% RSLogix 500 project MIXING.RSS, saved by version 8.30.00.16 %
PROJECT "UNTITLED"    % processor: MicroLogix 1000 %

PROGRAM FILES
  LAD 2 "MAIN_PROG"  6 rungs
  LAD 3 "USER_FAULT"  1 rungs
  LAD 4 "HSC_INT"  1 rungs
  LAD 5 "STI_INT"  1 rungs
  LAD 6, 7, 8, 9, 10, 11, 12, 13, 14, 15, 16: only END

DATA FILES
  O0 OUTPUT  5 elements
  I1 INPUT  8 elements
  S2 STATUS  33 elements
  B3 BINARY  32 elements
  T4 TIMER  40 elements
  C5 COUNTER  32 elements
  R6 CONTROL  16 elements
  N7 INTEGER  105 elements

LADDER 2 "MAIN_PROG"
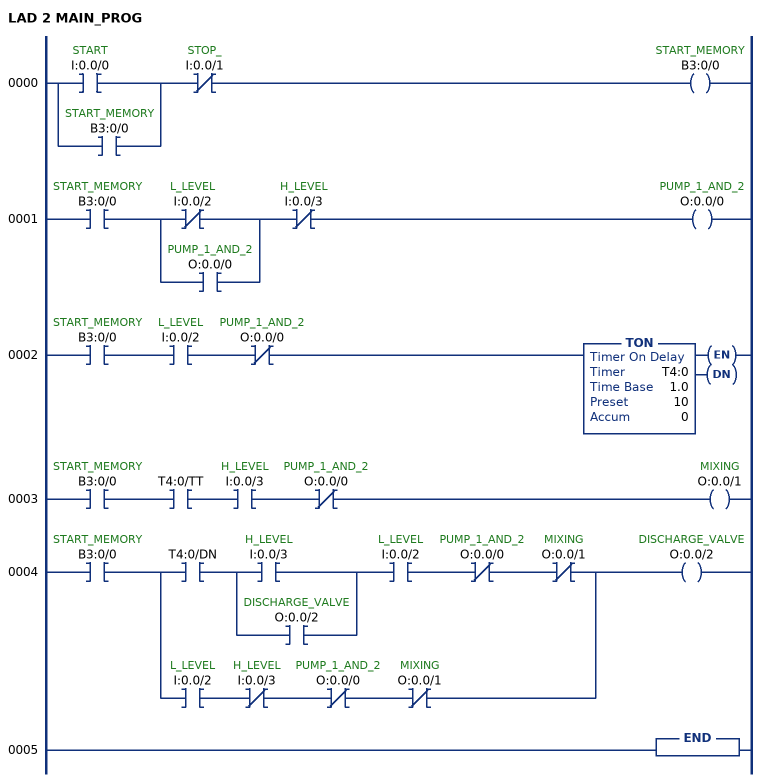
% Rung: 0 %
SOR BST XIC I:0.0/0 NXB XIC B3:0/0 BND XIO I:0.0/1 OTE B3:0/0 EOR
%   I:0.0/0  START %
%   B3:0/0  START_MEMORY %
%   I:0.0/1  STOP_ %
% Rung: 1 %
SOR XIC B3:0/0 BST XIO I:0.0/2 NXB XIC O:0.0/0 BND XIO I:0.0/3 OTE O:0.0/0 EOR
%   B3:0/0  START_MEMORY %
%   I:0.0/2  L_LEVEL %
%   O:0.0/0  PUMP_1_AND_2 %
%   I:0.0/3  H_LEVEL %
% Rung: 2 %
SOR XIC B3:0/0 XIC I:0.0/2 XIO O:0.0/0 TON T4:0 1.0 10 0 EOR
%   B3:0/0  START_MEMORY %
%   I:0.0/2  L_LEVEL %
%   O:0.0/0  PUMP_1_AND_2 %
% Rung: 3 %
SOR XIC B3:0/0 XIC T4:0/TT XIC I:0.0/3 XIO O:0.0/0 OTE O:0.0/1 EOR
%   B3:0/0  START_MEMORY %
%   I:0.0/3  H_LEVEL %
%   O:0.0/0  PUMP_1_AND_2 %
%   O:0.0/1  MIXING %
% Rung: 4 %
SOR XIC B3:0/0 BST XIC T4:0/DN BST XIC I:0.0/3 NXB XIC O:0.0/2 BND XIC I:0.0/2 XIO O:0.0/0 XIO O:0.0/1 NXB XIC I:0.0/2 XIO I:0.0/3 XIO O:0.0/0 XIO O:0.0/1 BND OTE O:0.0/2 EOR
%   B3:0/0  START_MEMORY %
%   I:0.0/3  H_LEVEL %
%   O:0.0/2  DISCHARGE_VALVE %
%   I:0.0/2  L_LEVEL %
%   O:0.0/0  PUMP_1_AND_2 %
%   O:0.0/1  MIXING %
% Rung: 5 %
SOR END EOR

DATA TABLE (non-zero values as saved)
DATA T4
% .PRE .ACC %
% T4:0 % 10 0
